// TIA Portal V19 export
DATA_BLOCK "Tacho2_EM06"   // DB7
VERSION : 1.0
// stored: InstanceOfName EM06_Descarga, InstanceOfType FB
"EM06_Descarga"
   // VAR_INPUT
   //    In : "EM06_Input";
   //    RecibidorLevelPV : Real;
   //    TachoLevelPV : Real;
   // END_VAR
   // VAR_OUTPUT
   //    Out : "EM06_Output";
   //    CM_Vlv_Descarga_Out : Bool;
   //    CM_Vlv_Desague_Out : Bool;
   //    CMAlarm : Bool;
   // END_VAR
   // VAR
   //    State : Int;
   //    ActiveMode : Int;
   //    DrainElapsed : Time;
   //    AlarmLatched : Bool;
   //    FaultCode : Int;
   //    TimerEmpty { S7_SetPoint := 'True'} : TON_TIME;
   //    TimerDrain { S7_SetPoint := 'True'} : TON_TIME;
   //    TrigStart { S7_SetPoint := 'True'} : R_TRIG;
   //    TrigStop { S7_SetPoint := 'True'} : R_TRIG;
   //    TrigHold { S7_SetPoint := 'True'} : R_TRIG;
   //    TrigAbort { S7_SetPoint := 'True'} : R_TRIG;
   //    TrigReset { S7_SetPoint := 'True'} : R_TRIG;
   //    CM_Vlv_Descarga { S7_SetPoint := 'True'} : "VlvL";
   //    CM_Vlv_Desague { S7_SetPoint := 'True'} : "VlvL";
   // END_VAR
BEGIN
END_DATA_BLOCK
